(* IEC 61131-3 sources: POMIRTS_lab3/AS/Library_2/AsSafety, 3 files *)

(* ---- AsSafety.fun ---- *)
{REDUND_ERROR} FUNCTION_BLOCK safeRemoteControl (*Remote Control Function Block*)
	VAR_INPUT
		SafeLOGICID : UINT; (*SafeLOGIC ID*)
		Execute : BOOL; (*execution*)
		pCommandData : UDINT; (*pointer to command data*)
	END_VAR
	VAR_OUTPUT
		Done : BOOL; (*execution done*)
		Busy : BOOL; (*execution busy*)
		Error : BOOL; (*execution error*)
		StatusID : UINT; (*execution status: ERR_OK, ERR_FUB_BUSY, 0xXXXX = see help*)
		SafeLOGICStatus : RemoteControlStatusTypeV1; (*SafeLOGIC status*)
	END_VAR
	VAR
		i_state : UINT; (*internal variable*)
		i_result : UINT; (*internal variable*)
		i_tmp : UDINT; (*internal variable*)
		i_handle : UDINT; (*internal variable*)
	END_VAR
END_FUNCTION_BLOCK

{REDUND_ERROR} FUNCTION_BLOCK safeRemoteControl_V2 (*Remote Control Function Block*)
	VAR_INPUT
		SafeLOGICID : UINT; (*SafeLOGIC ID*)
		Execute : BOOL; (*execution*)
		pCommandData : UDINT; (*pointer to command data*)
	END_VAR
	VAR_OUTPUT
		Done : BOOL; (*execution done*)
		Busy : BOOL; (*execution busy*)
		Error : BOOL; (*execution error*)
		StatusID : UINT; (*execution status: ERR_OK, ERR_FUB_BUSY, 0xXXXX = see help*)
		SafeLOGICStatus : RemoteControlStatusTypeV2; (*SafeLOGIC status*)
	END_VAR
	VAR
		Internal : AsSafetyInternalType; (*internal variable*)
	END_VAR
END_FUNCTION_BLOCK

{REDUND_ERROR} FUNCTION_BLOCK safeDownloadApplication (*Download Application Function Block*)
	VAR_INPUT
		SafeLOGICID : UINT; (*SafeLOGIC ID*)
		Execute : BOOL; (*execution*)
		pCommandData : UDINT; (*pointer to command data*)
	END_VAR
	VAR_OUTPUT
		Done : BOOL; (*execution done*)
		Busy : BOOL; (*execution busy*)
		Error : BOOL; (*execution error*)
		StatusID : UINT; (*execution status: ERR_OK, ERR_FUB_BUSY, 0xXXXX = see help*)
		UnlockRequired : BOOL; (*unlock required*)
		ApplicationCRC : UDINT; (*application CRC*)
	END_VAR
	VAR
		i_state : UINT; (*internal variable*)
		i_result : UINT; (*internal variable*)
		i_tmp : UDINT; (*internal variable*)
		i_handle : UDINT; (*internal variable*)
	END_VAR
END_FUNCTION_BLOCK

{REDUND_ERROR} FUNCTION_BLOCK safeDownloadApplication_V2 (*Download Application Function Block*)
	VAR_INPUT
		SafeLOGICID : UINT; (*SafeLOGIC ID*)
		Execute : BOOL; (*execution*)
		pCommandData : UDINT; (*pointer to command data*)
	END_VAR
	VAR_OUTPUT
		Done : BOOL; (*execution done*)
		Busy : BOOL; (*execution busy*)
		Error : BOOL; (*execution error*)
		StatusID : UINT; (*execution status: ERR_OK, ERR_FUB_BUSY, 0xXXXX = see help*)
		UnlockRequired : BOOL; (*unlock required*)
		ApplicationCRC : UDINT; (*application CRC*)
	END_VAR
	VAR
		Internal : AsSafetyInternalType; (*internal variable*)
	END_VAR
END_FUNCTION_BLOCK

{REDUND_ERROR} FUNCTION_BLOCK safeDownloadData (*Download Data Function Block*)
	VAR_INPUT
		SafeLOGICID : UINT; (*SafeLOGIC ID*)
		Execute : BOOL; (*execution*)
		Type : UINT; (*type of data: safeDATA_TYPE_MAOP, safeDATA_TYPE_EXTMAOP,... *)
		pCommandData : UDINT; (*pointer to command data*)
	END_VAR
	VAR_OUTPUT
		Done : BOOL; (*execution done*)
		Busy : BOOL; (*execution busy*)
		Error : BOOL; (*execution error*)
		StatusID : UINT; (*execution status: ERR_OK, ERR_FUB_BUSY, 0xXXXX = see help*)
		UnlockRequired : BOOL; (*unlock required*)
		Timestamp : UDINT; (*timestamp from data*)
	END_VAR
	VAR
		i_state : UINT; (*internal variable*)
		i_result : UINT; (*internal variable*)
		i_tmp : UDINT; (*internal variable*)
		i_handle : UDINT; (*internal variable*)
	END_VAR
END_FUNCTION_BLOCK

{REDUND_ERROR} FUNCTION_BLOCK safeDownloadData_V2 (*Download Data Function Block*)
	VAR_INPUT
		SafeLOGICID : UINT; (*SafeLOGIC ID*)
		Execute : BOOL; (*execution*)
		Type : UINT; (*type of data: safeDATA_TYPE_MAOP, safeDATA_TYPE_EXTMAOP,... *)
		pCommandData : UDINT; (*pointer to command data*)
	END_VAR
	VAR_OUTPUT
		Done : BOOL; (*execution done*)
		Busy : BOOL; (*execution busy*)
		Error : BOOL; (*execution error*)
		StatusID : UINT; (*execution status: ERR_OK, ERR_FUB_BUSY, 0xXXXX = see help*)
		UnlockRequired : BOOL; (*unlock required*)
		Timestamp : UDINT; (*timestamp from data*)
	END_VAR
	VAR
		Internal : AsSafetyInternalType; (*internal variable*)
	END_VAR
END_FUNCTION_BLOCK

{REDUND_ERROR} FUNCTION_BLOCK safeConfigurationOnTarget (*Configuration On Target Function Block*)
	VAR_INPUT
		SafeLOGICID : UINT; (*SafeLOGIC ID*)
		Execute : BOOL; (*execution*)
		Type : UINT; (*type of data: safeDATA_TYPE_MAOP, safeDATA_TYPE_EXTMAOP,...*)
		pCommandData : UDINT; (*pointer to command data*)
	END_VAR
	VAR_OUTPUT
		Done : BOOL; (*execution done*)
		Busy : BOOL; (*execution busy*)
		Error : BOOL; (*execution error*)
		StatusID : UINT; (*execution status: ERR_OK, ERR_FUB_BUSY, 0xXXXX = see help*)
		Timestamp : UDINT; (*timestamp of data*)
	END_VAR
	VAR
		i_state : UINT; (*internal variable*)
		i_result : UINT; (*internal variable*)
		i_tmp : UDINT; (*internal variable*)
		i_handle : UDINT; (*internal variable*)
	END_VAR
END_FUNCTION_BLOCK

{REDUND_ERROR} FUNCTION_BLOCK safeConfigurationOnTarget_V2 (*Configuration On Target Function Block*)
	VAR_INPUT
		SafeLOGICID : UINT; (*SafeLOGIC ID*)
		Execute : BOOL; (*execution*)
		Type : UINT; (*type of data: safeDATA_TYPE_MAOP, safeDATA_TYPE_EXTMAOP,...*)
		pCommandData : UDINT; (*pointer to command data*)
	END_VAR
	VAR_OUTPUT
		Done : BOOL; (*execution done*)
		Busy : BOOL; (*execution busy*)
		Error : BOOL; (*execution error*)
		StatusID : UINT; (*execution status: ERR_OK, ERR_FUB_BUSY, 0xXXXX = see help*)
		Timestamp : UDINT; (*timestamp of data*)
	END_VAR
	VAR
		Internal : AsSafetyInternalType; (*internal variable*)
	END_VAR
END_FUNCTION_BLOCK

{REDUND_ERROR} FUNCTION safeLibraryVersion : UINT (*returns the actual library version*)
END_FUNCTION

{REDUND_ERROR} FUNCTION_BLOCK safeDownloadFile (*Download File Function Block*)
	VAR_INPUT
		SafeLOGICID : UINT; (*SafeLOGIC ID*)
		Execute : BOOL; (*execution*)
		pCommandData : UDINT; (*pointer to command data*)
	END_VAR
	VAR_OUTPUT
		Done : BOOL; (*execution done*)
		Busy : BOOL; (*execution busy*)
		Error : BOOL; (*execution error*)
		StatusID : UINT; (*execution status: ERR_OK, ERR_FUB_BUSY, 0xXXXX = see help*)
		UnlockRequired : BOOL; (*unlock required*)
		Timestamp : UDINT; (*timestamp from data*)
	END_VAR
	VAR
		Internal : AsSafetyInternalType; (*internal variable*)
	END_VAR
END_FUNCTION_BLOCK

{REDUND_ERROR} FUNCTION_BLOCK safeCheckTable (*Check Table Function Block*)
	VAR_INPUT
		Execute : BOOL; (*execution*)
		InstNr : USINT; (*instance number*)
		pUser : UDINT; (*user name*)
		Timestamp : UDINT; (*timestamp*)
		TableType : USINT; (*table type*)
		EntryCnt : UDINT; (*number of entries*)
		pTableHeader : UDINT; (*table header input*)
		pTableData : UDINT; (*table data input*)
		pTableHeaderOut : UDINT; (*table header output buffer*)
		pTableDataOut : UDINT; (*table data output buffer*)
		pFileDataOut : UDINT; (*file data output buffer*)
		AckData : USINT; (*1 .. acknowledge table data, 2 .. NOT acknowledge table data, abort FUB*)
	END_VAR
	VAR_OUTPUT
		Done : BOOL; (*execution done*)
		Busy : BOOL; (*execution busy*)
		Error : BOOL; (*execution error*)
		StatusID : UINT; (*execution status: ERR_OK, ERR_FUB_BUSY, 0xXXXX = see help*)
		CheckErrorCode : UDINT; (*table check error code*)
		CheckErrorLine : UDINT; (*table check error line*)
		CheckErrorColumn : UDINT; (*table check error column*)
		pCrcOut : UDINT; (*returns pointer to CRC data*)
		CrcCntOut : UDINT; (*returns number of CRCs*)
	END_VAR
	VAR
		i_step : UINT; (*internal*)
		i_tmp : UDINT; (*internal*)
		i_clean : BOOL; (*internal*)
	END_VAR
END_FUNCTION_BLOCK

{REDUND_ERROR} FUNCTION_BLOCK safeFileInfo (*File Info Function Block*)
	VAR_INPUT
		SafeLOGICID : UINT; (*SafeLOGIC ID*)
		Execute : BOOL; (*execution*)
		Type : UINT; (*type of data: safeDATA_TYPE_MAOP, safeDATA_TYPE_EXTMAOP,...*)
		pCommandData : UDINT; (*pointer to command data*)
	END_VAR
	VAR_OUTPUT
		Done : BOOL; (*execution done*)
		Busy : BOOL; (*execution busy*)
		Error : BOOL; (*execution error*)
		StatusID : UINT; (*execution status: ERR_OK, ERR_FUB_BUSY, 0xXXXX = see help*)
	END_VAR
	VAR
		Internal : AsSafetyInternalType; (*internal variable*)
	END_VAR
END_FUNCTION_BLOCK

{REDUND_ERROR} FUNCTION safeGetTableLength : UDINT (*Function returns size of table data*)
	VAR_INPUT
		TableType : USINT; (*table type*)
		EntryCnt : UDINT; (*number of entries*)
		pTableHeader : UDINT; (*pointer to table header*)
	END_VAR
END_FUNCTION

{REDUND_ERROR} FUNCTION_BLOCK safeGetDataLength (*Function Block returns size of download file*)
	VAR_INPUT
		Execute : BOOL; (*execution*)
		Type : UINT; (*type of data: safeDATA_TYPE_MAOP, safeDATA_TYPE_EXTMAOP,... *)
		pCommandData : UDINT; (*pointer to command data*)
	END_VAR
	VAR_OUTPUT
		Done : BOOL; (*execution done*)
		Busy : BOOL; (*execution busy*)
		Error : BOOL; (*execution error*)
		StatusID : UINT; (*execution status: ERR_OK, ERR_FUB_BUSY, 0xXXXX = see help*)
		Length : UDINT; (*calculated length of download file*)
	END_VAR
	VAR
		Internal : AsSafetyInternalType; (*internal variable*)
	END_VAR
END_FUNCTION_BLOCK

{REDUND_ERROR} FUNCTION_BLOCK safeCreateData (*Create Data Function Block*)
	VAR_INPUT
		SafeLOGICID : UINT; (*SafeLOGIC ID*)
		Execute : BOOL; (*execution*)
		Type : UINT; (*type of data: safeDATA_TYPE_MAOP, safeDATA_TYPE_EXTMAOP,... *)
		pCommandData : UDINT; (*pointer to command data*)
		FileDataOutLen : UDINT; (*size of buffer for file data*)
		pFileDataOut : UDINT; (*pointer to memory buffer for file data*)
	END_VAR
	VAR_OUTPUT
		Done : BOOL; (*execution done*)
		Busy : BOOL; (*execution busy*)
		Error : BOOL; (*execution error*)
		StatusID : UINT; (*execution status: ERR_OK, ERR_FUB_BUSY, 0xXXXX = see help*)
		UnlockRequired : BOOL; (*unlock required*)
		Timestamp : UDINT; (*timestamp from data*)
	END_VAR
	VAR
		Internal : AsSafetyInternalType; (*internal variable*)
	END_VAR
END_FUNCTION_BLOCK

{REDUND_ERROR} FUNCTION_BLOCK safeLogicInfo (*Remote Control Function Block*)
	VAR_INPUT
		SafeLOGICID : UINT; (*SafeLOGIC ID*)
		Execute : BOOL; (*execution*)
		Type : UINT; (*type of data: safeINFO_TYPE_PWD_INFO, safeINFO_TYPE_PWD_CHK, safeINFO_TYPE_UDID_INFO*)
		pCommandData : UDINT; (*pointer to command data*)
	END_VAR
	VAR_OUTPUT
		Done : BOOL; (*execution done*)
		Busy : BOOL; (*execution busy*)
		Error : BOOL; (*execution error*)
		StatusID : UINT; (*execution status: ERR_OK, ERR_FUB_BUSY, 0xXXXX = see help*)
	END_VAR
	VAR
		Internal : AsSafetyInternalType; (*internal variable*)
	END_VAR
END_FUNCTION_BLOCK

(* ---- AsSafety.typ ---- *)
TYPE
	FileReferenceType : 	STRUCT  (*file reference*)
		Device : STRING[80]; (*pointer to the device name*)
		File : STRING[80]; (*pointer to the file name*)
	END_STRUCT;
	AsSafetyInternalType : 	STRUCT  (*internal data type*)
		Clean : BOOL;
		State : UINT;
		Result : UINT;
		Tmp : UDINT;
		pThis : UDINT;
		pFcn : UDINT;
	END_STRUCT;
	SourceLocalDataTypeV1 : 	STRUCT  (*local data source type*)
		pFileData : UDINT; (*pointer to data buffer*)
		FileLength : UDINT; (*data length*)
	END_STRUCT;
	SourceLocalFileTypeV1 : 	STRUCT  (*local file source*)
		SourceFile : FileReferenceType; (*path to local file*)
	END_STRUCT;
	DataSourceTypeV1 : 	STRUCT  (*source data type*)
		Type : UINT; (*0 .. file upload from safeLOGIC, 1 .. local data buffer, 2 .. local file*)
		LocalData : SourceLocalDataTypeV1; (*arguments for local data*)
		LocalFile : SourceLocalFileTypeV1; (*arguments for local file*)
	END_STRUCT;
	InfoCmdPwdInfoTypeV1 : 	STRUCT  (*password info data from SafeLOGIC command structure*)
		Version : UINT; (*used version*)
		PasswordSet : BOOL; (*0 .. no password set, 1 .. password is set*)
	END_STRUCT;
	InfoCmdPwdChkTypeV1 : 	STRUCT  (*password check data from SafeLOGIC command structure*)
		Version : UINT; (*used version*)
		Password : STRING[16]; (*password for check*)
		PasswordEqual : BOOL; (*0 .. no password set, 1 .. password is set*)
	END_STRUCT;
	ConfigurationAddParaTypeV2 : 	STRUCT  (*additional parameter data from SafeLOGIC*)
		SADR : UINT; (*safety address*)
		ID : USINT; (*id*)
		pParaData : UDINT; (*pointer to additional parameter data*)
		Length : UDINT; (*size of parameter buffer*)
		LengthOut : UDINT; (*length of parameter*)
		CRC : UDINT; (*CRC*)
		Timestamp : UDINT; (*timestamp*)
	END_STRUCT;
	ConfigurationAddParaTypeV1 : 	STRUCT  (*additional parameter data from SafeLOGIC*)
		SADR : UINT; (*safety address*)
		ID : USINT; (*id*)
		pParaData : UDINT; (*pointer to additional parameter data*)
		Length : UDINT; (*size of parameter buffer*)
		CRC : UDINT; (*CRC*)
		Timestamp : UDINT; (*timestamp*)
	END_STRUCT;
	ConfigurationBitOptionsTypeV1 : 	STRUCT  (*bit machine options*)
		BitData : ARRAY[0..63]OF USINT; (*bit array*)
	END_STRUCT;
	ConfigurationCmdAddParaTypeV2 : 	STRUCT  (*additional parameter data from SafeLOGIC command structure*)
		Version : UINT; (*input data: used version*)
		Password : STRING[16]; (*input data: password*)
		pParaDataOutput : UDINT; (*input data: pointer to list of type ConfigurationAddParaTypeV2*)
		NumberParaSetsOutput : UINT; (*input data: number of available entries in pParaDataOutput*)
		NumberParaSetsOutputOut : UINT; (*return value: number of returned entries*)
		pBackupFile : UDINT; (*input data: 0 .. no backup, otherwise pointer to struct of type FileReferenceType *)
		pXmlOutputFile : UDINT; (*input data: 0 .. don't create XML output data, otherwise pointer to struct of type FileReferenceType*)
	END_STRUCT;
	ConfigurationCmdAddParaTypeV1 : 	STRUCT  (*additional parameter data from SafeLOGIC command structure*)
		Version : UINT; (*input data: used version*)
		Password : STRING[16]; (*input data: password*)
		pParaDataOutput : UDINT; (*return value: pointer to list of type ConfigurationAddParaTypeV1*)
		NumberParaSetsOutput : UINT; (*return value: number of returned entries*)
	END_STRUCT;
	ConfigurationCmdExtMaOpTypeV2 : 	STRUCT  (*extended machine options from SafeLOGIC command structure*)
		Version : UINT; (*input data: safeVERSION_R110*)
		Password : STRING[16]; (*input data: password*)
		pIntDataOutput : UDINT; (*input data: pointer to list of type ConfigurationIntOptionsTypeV1*)
		NumberIntOutput : UINT; (*input data: number of available entries in INT buffer*)
		NumberIntOutputOut : UINT; (*return value: number of returned INT data entries*)
		pUintDataOutput : UDINT; (*input data: pointer to list of type ConfigurationUintOptionsTypeV1*)
		NumberUintOutput : UINT; (*input data: number of available entries in UINT buffer*)
		NumberUintOutputOut : UINT; (*return value: number of returned UINT data entries*)
		pDintDataOutput : UDINT; (*input data: pointer to list of type ConfigurationDintOptionsTypeV1*)
		NumberDintOutput : UINT; (*input data: number of available DINT data entries*)
		NumberDintOutputOut : UINT; (*return value: number of returned DINT data entries*)
		pUdintDataOutput : UDINT; (*input data: pointer to list of type ConfigurationUdintOptionsTypeV1*)
		NumberUdintOutput : UINT; (*input data: number of available UDINT data entries*)
		NumberUdintOutputOut : UINT; (*return value: number of returned UDINT data entries*)
		pBackupFile : UDINT; (*input data: 0 .. no backup, otherwise pointer to struct of type FileReferenceType *)
		pXmlOutputFile : UDINT; (*input data: 0 .. don't create XML output data, otherwise pointer to struct of type FileReferenceType*)
	END_STRUCT;
	ConfigurationCmdExtMaOpTypeV1 : 	STRUCT  (*extended machine options from SafeLOGIC command structure*)
		Version : UINT; (*input data: safeVERSION_R107*)
		Password : STRING[16]; (*input data: password*)
		pIntDataOutput : UDINT; (*return value: pointer to list of type ConfigurationIntOptionsTypeV1*)
		NumberIntOutput : UINT; (*return value: number of returned INT data entries*)
		pUintDataOutput : UDINT; (*return value: pointer to list of type ConfigurationUintOptionsTypeV1*)
		NumberUintOutput : UINT; (*return value: number of returned UINT data entries*)
		pDintDataOutput : UDINT; (*return value: pointer to list of type ConfigurationDintOptionsTypeV1*)
		NumberDintOutput : UINT; (*return value: number of returned DINT data entries*)
		pUdintDataOutput : UDINT; (*return value: pointer to list of type ConfigurationUdintOptionsTypeV1*)
		NumberUdintOutput : UINT; (*return value: number of returned UDINT data entries*)
	END_STRUCT;
	ConfigurationCmdMaOpTypeV2 : 	STRUCT  (*machine options from SafeLOGIC command structure Version 2*)
		Version : UINT; (*input data: safeVERSION_R110*)
		Password : STRING[16]; (*input data: password*)
		pDeviceListOutput : UDINT; (*input data: pointer to device list buffer of type ConfigurationDeviceTypeV1*)
		NumberDevicesOutput : UINT; (*input data: number of available device entries in devices list buffer*)
		NumberDevicesOutputOut : UINT; (*return value: number of returned device entries*)
		pMachineOptionsOutput : UDINT; (*input data: pointer to bit machine options of type ConfigurationBitOptionsTypeV1*)
		pModuleFlagsOutput : UDINT; (*input data: pointer to module flags of type ConfigurationModuleFlagsTypeV1*)
		pBackupFile : UDINT; (*input data: 0 .. no backup, otherwise pointer to struct of type FileReferenceType *)
		pXmlOutputFile : UDINT; (*input data: 0 .. don't create XML output data, otherwise pointer to struct of type FileReferenceType*)
	END_STRUCT;
	ConfigurationCmdMaOpTypeV1 : 	STRUCT  (*machine options from SafeLOGIC command structure Version 1*)
		Version : UINT; (*input data: safeVERSION_R107*)
		Password : STRING[16]; (*input data: password*)
		pDeviceListOutput : UDINT; (*return value: pointer to device list of type ConfigurationDeviceTypeV1*)
		NumberDevicesOutput : UINT; (*return value: number of returned entries*)
		pMachineOptionsOutput : UDINT; (*return value: pointer to bit machine options of type ConfigurationBitOptionsTypeV1*)
		pModuleFlagsOutput : UDINT; (*return value: pointer to module flags of type ConfigurationModuleFlagsTypeV1*)
	END_STRUCT;
	ConfigurationCmdTableTypeV2 : 	STRUCT  (*table data from SafeLOGIC command structure*)
		Version : UINT; (*input data: safeVERSION_R110*)
		Password : STRING[16]; (*input data: password*)
		pTableDataOutput : UDINT; (*input data: pointer to list of type ConfigurationTableTypeV1*)
		NumberTablesOutput : UINT; (*input data: number of available entries in pTableDataOutput*)
		NumberTablesOutputOut : UINT; (*return value: number of returned table entries*)
		pBackupFile : UDINT; (*input data: 0 .. no backup, otherwise pointer to struct of type FileReferenceType *)
		pXmlOutputFile : UDINT; (*input data: 0 .. don't create XML output data, otherwise pointer to struct of type FileReferenceType*)
	END_STRUCT;
	ConfigurationCmdTableTypeV1 : 	STRUCT  (*table data from SafeLOGIC command structure*)
		Version : UINT; (*input data: safeVERSION_R107*)
		Password : STRING[16]; (*input data: password*)
		pTableDataOutput : UDINT; (*return value: pointer to list of type ConfigurationTableTypeV1*)
		NumberTablesOutput : UINT; (*return value: number of returned table entries*)
	END_STRUCT;
	FileInfoCmdTypeV1 : 	STRUCT  (*file info command structure*)
		Version : UINT; (*used version*)
		DataSource : DataSourceTypeV1; (*data source*)
		Timestamp : UDINT; (*timestamp*)
		pCrcs : UDINT; (*buffer for CRCs*)
		NumberOfCrcs : UINT; (*size of CRC buffer*)
		NumberOfCrcsOut : UINT; (*number of CRCs*)
	END_STRUCT;
	ConfigurationDeviceTypeV1 : 	STRUCT  (*safety device from SafeLOGIC*)
		SADR : UINT; (*safety address*)
		UDID : ARRAY[0..5]OF USINT; (*UDID*)
	END_STRUCT;
	ConfigurationDintOptionsTypeV1 : 	STRUCT  (*DINT machine options*)
		ID : UINT; (*id*)
		Value : DINT; (*value*)
	END_STRUCT;
	ConfigurationIntOptionsTypeV1 : 	STRUCT  (*INT machine options*)
		ID : UINT; (*id*)
		Value : INT; (*value*)
	END_STRUCT;
	ConfigurationModuleFlagsTypeV1 : 	STRUCT  (*module flags*)
		Optional : ARRAY[0..127]OF USINT; (*optional*)
		Startup : ARRAY[0..127]OF USINT; (*startup*)
		NotPresent : ARRAY[0..127]OF USINT; (*not present*)
	END_STRUCT;
	ConfigurationTableTypeV2 : 	STRUCT  (*table data for command struct V1*)
		ID : UINT; (*table id*)
		Type : USINT; (*table type*)
		NumberOfCRCs : UINT; (*input data: number of available entries in pCRCData*)
		NumberOfCRCsOut : UINT; (*return value: number of returned CRC entries*)
		pCRCData : UDINT; (*input data: pointer to table CRC buffer*)
	END_STRUCT;
	ConfigurationTableTypeV1 : 	STRUCT  (*table data for command struct V2*)
		ID : UINT; (*table id*)
		Type : USINT; (*table type*)
		NumberOfCRCs : UINT; (*return value: number of returned CRCs*)
		pCRCData : UDINT; (*return value: pointer to table CRC buffer*)
	END_STRUCT;
	ConfigurationUdintOptionsTypeV1 : 	STRUCT  (*UDINT machine options*)
		ID : UINT; (*id*)
		Value : UDINT; (*value*)
	END_STRUCT;
	ConfigurationUintOptionsTypeV1 : 	STRUCT  (*UINT machine options*)
		ID : UINT; (*id*)
		Value : UINT; (*value*)
	END_STRUCT;
	DownloadAcknExtMaOpTypeV1 : 	STRUCT  (*acknowledge extended machine options structure*)
		AcknIntOptions : ARRAY[0..63]OF BOOL; (*acknowledge INT*)
		AcknUintOptions : ARRAY[0..63]OF BOOL; (*acknowledge UINT*)
		AcknDintOptions : ARRAY[0..63]OF BOOL; (*acknowledge DINT*)
		AcknUdintOptions : ARRAY[0..63]OF BOOL; (*acknowledge UDINT*)
	END_STRUCT;
	DownloadAcknMaOpTypeV1 : 	STRUCT  (*acknowledge bit machine options structure*)
		AcknBitOptions : ARRAY[0..63]OF USINT; (*acknowledge bit*)
	END_STRUCT;
	DownloadAcknAddParaTypeV1 : 	STRUCT  (*acknowledge bit additional parameter*)
		AcknBitAddPara : ARRAY[0..63]OF USINT; (*acknowledge bit*)
	END_STRUCT;
	DownloadCmdAddParaTypeV2 : 	STRUCT  (*additional paramater command structure*)
		Version : UINT; (*input data: used version*)
		Password : STRING[16]; (*input data: password*)
		UDID_Low : UDINT; (*input data: UDID low*)
		UDID_High : UINT; (*input data: UDID high*)
		Unlock : USINT; (*input data: unlock data*)
		pParaListInput : UDINT; (*input data: pointer to additional parameter input data list of type DownloadAddParaTypeV1*)
		NumberParaSetsInput : UINT; (*input data: number of input parameter entries in pParaListInput*)
		pParaDataOutput : UDINT; (*input data: pointer to list of type ConfigurationAddParaTypeV2*)
		NumberParaSetsOutput : UINT; (*input data: number of available entries in pParaDataOutput*)
		NumberParaSetsOutputOut : UINT; (*return value: number of returned entries*)
		pBackupFile : UDINT; (*input data: 0 .. no backup, otherwise pointer to struct of type FileReferenceType *)
		pXmlOutputFile : UDINT; (*input data: 0 .. don't create XML output data, otherwise pointer to struct of type FileReferenceType*)
	END_STRUCT;
	DownloadCmdAddParaTypeV1 : 	STRUCT  (*additional paramater command structure*)
		Version : UINT; (*input data: used version*)
		Password : STRING[16]; (*input data: password*)
		UDID_Low : UDINT; (*input data: UDID low*)
		UDID_High : UINT; (*input data: UDID high*)
		Unlock : USINT; (*input data: unlock data*)
		pParaListInput : UDINT; (*input data: pointer to additional parameter input data list of type DownloadAddParaTypeV1*)
		NumberParaSetsInput : UINT; (*input data: number of input parameter entries in pParaListInput*)
		pParaDataOutput : UDINT; (*return value: pointer to list of type ConfigurationAddParaTypeV1*)
		NumberParaSetsOutput : UINT; (*return value: number of returned entries*)
	END_STRUCT;
	DownloadCmdApplicationTypeV1 : 	STRUCT  (*application command structure*)
		Version : UINT; (*used version*)
		Password : STRING[16]; (*password*)
		UDID_Low : UDINT; (*UDID low*)
		UDID_High : UINT; (*UDID high*)
		ApplicationID : UINT; (*application id*)
		Device : STRING[80]; (*device for file*)
		File : STRING[80]; (*file name*)
		Unlock : USINT; (*unlock application*)
	END_STRUCT;
	DownloadCmdExtMaOpTypeV2 : 	STRUCT  (*extended machine options command structure*)
		Version : UINT; (*input data: safeVERSION_R110*)
		Password : STRING[16]; (*input data: password*)
		UDID_Low : UDINT; (*input data: UDID low*)
		UDID_High : UINT; (*input data: UDID high*)
		Unlock : USINT; (*input data: unlock data*)
		pIntDataInput : UDINT; (*input data: pointer to INT input data list from type ConfigurationIntOptionsTypeV1*)
		NumberIntInput : UINT; (*input data: number of INT input entries in pIntDataInput*)
		pUintDataInput : UDINT; (*input data: pointer to UINT input data list from type ConfigurationUintOptionsTypeV1*)
		NumberUintInput : UINT; (*input data: number of UINT input entries in pUintDataInput*)
		pDintDataInput : UDINT; (*input data: pointer to DINT input data list from type ConfigurationDintOptionsTypeV1*)
		NumberDintInput : UINT; (*input data: number of DINT input entries in pDintDataInput*)
		pUdintDataInput : UDINT; (*input data: pointer to UDINT input data list from type ConfigurationUdintOptionsTypeV1*)
		NumberUdintInput : UINT; (*input data: number of UDINT input entries in pUdintDataInput*)
		pAcknMachineOptions : UDINT; (*input data: pointer to acknowledge information of type DownloadAcknMaOpTypeV1*)
		pIntDataOutput : UDINT; (*input data: pointer to list of type ConfigurationIntOptionsTypeV1*)
		NumberIntOutput : UINT; (*input data: number of available entries in INT buffer*)
		NumberIntOutputOut : UINT; (*return value: number of returned INT data entries*)
		pUintDataOutput : UDINT; (*input data: pointer to list of type ConfigurationUintOptionsTypeV1*)
		NumberUintOutput : UINT; (*input data: number of available entries in UINT buffer*)
		NumberUintOutputOut : UINT; (*return value: number of returned UINT data entries*)
		pDintDataOutput : UDINT; (*input data: pointer to list of type ConfigurationDintOptionsTypeV1*)
		NumberDintOutput : UINT; (*input data: number of available DINT data entries*)
		NumberDintOutputOut : UINT; (*return value: number of returned DINT data entries*)
		pUdintDataOutput : UDINT; (*input data: pointer to list of type ConfigurationUdintOptionsTypeV1*)
		NumberUdintOutput : UINT; (*input data: number of available UDINT data entries*)
		NumberUdintOutputOut : UINT; (*number of UDINT channels from SafeLOGIC*)
		pBackupFile : UDINT; (*input data: 0 .. no backup, otherwise pointer to struct of type FileReferenceType *)
		pXmlOutputFile : UDINT; (*input data: 0 .. don't create XML output data, otherwise pointer to struct of type FileReferenceType*)
	END_STRUCT;
	DownloadCmdExtMaOpTypeV1 : 	STRUCT  (*return value: number of returned UDINT data entries*)
		Version : UINT; (*input data: safeVERSION_R107*)
		Password : STRING[16]; (*input data: password*)
		UDID_Low : UDINT; (*input data: UDID low*)
		UDID_High : UINT; (*input data: UDID high*)
		Unlock : USINT; (*input data: unlock data*)
		pIntDataInput : UDINT; (*input data: pointer to INT input data list from type ConfigurationIntOptionsTypeV1*)
		NumberIntInput : UINT; (*input data: number of INT input entries in pIntDataInput*)
		pUintDataInput : UDINT; (*input data: pointer to UINT input data list from type ConfigurationUintOptionsTypeV1*)
		NumberUintInput : UINT; (*input data: number of UINT input entries in pUintDataInput*)
		pDintDataInput : UDINT; (*input data: pointer to DINT input data list from type ConfigurationDintOptionsTypeV1*)
		NumberDintInput : UINT; (*input data: number of DINT input entries in pDintDataInput*)
		pUdintDataInput : UDINT; (*input data: pointer to UDINT input data list from type ConfigurationUdintOptionsTypeV1*)
		NumberUdintInput : UINT; (*input data: number of UDINT input entries in pUdintDataInput*)
		pAcknMachineOptions : UDINT; (*input data: pointer to acknowledge information of type DownloadAcknMaOpTypeV1*)
		pIntDataOutput : UDINT; (*return value: pointer to list of type ConfigurationIntOptionsTypeV1*)
		NumberIntOutput : UINT; (*return value: number of returned INT data entries*)
		pUintDataOutput : UDINT; (*return value: pointer to list of type ConfigurationUintOptionsTypeV1*)
		NumberUintOutput : UINT; (*return value: number of returned UINT data entries*)
		pDintDataOutput : UDINT; (*return value: pointer to list of type ConfigurationDintOptionsTypeV1*)
		NumberDintOutput : UINT; (*return value: number of returned DINT data entries*)
		pUdintDataOutput : UDINT; (*return value: pointer to list of type ConfigurationUdintOptionsTypeV1*)
		NumberUdintOutput : UINT; (*return value: number of returned UDINT data entries*)
	END_STRUCT;
	DownloadCmdMaOpTypeV2 : 	STRUCT  (*machine options command structure*)
		Version : UINT; (*input data: safeVERSION_R110*)
		Password : STRING[16]; (*input data: password*)
		UDID_Low : UDINT; (*input data: UDID low from SafeLOGIC*)
		UDID_High : UINT; (*input data: UDID high from SafeLOGIC*)
		Unlock : USINT; (*input data: unlock data*)
		pDeviceListInput : UDINT; (*input data: pointer to input device list of type DownloadDeviceTypeV1*)
		NumberDevicesInput : UINT; (*input data: number of input devices*)
		pMachineOptionsInput : UDINT; (*input data: pointer to input bit machine options of type ConfigurationBitOptionsTypeV1*)
		pModuleFlagsInput : UDINT; (*input data: pointer to input module flags of type ConfigurationModuleFlagsTypeV1*)
		pAcknMachineOptions : UDINT; (*input data: pointer to acknowledge information of type DownloadAcknMaOpTypeV1*)
		pDeviceListOutput : UDINT; (*input data: pointer to device list buffer of type ConfigurationDeviceTypeV1*)
		NumberDevicesOutput : UINT; (*input data: number of available device entries in devices list buffer*)
		NumberDevicesOutputOut : UINT; (*return value: number of returned device entries*)
		pMachineOptionsOutput : UDINT; (*input data: pointer to bit machine options of type ConfigurationBitOptionsTypeV1*)
		pModuleFlagsOutput : UDINT; (*input data: pointer to module flags of type ConfigurationModuleFlagsTypeV1*)
		pBackupFile : UDINT; (*input data: 0 .. no backup, otherwise pointer to struct of type FileReferenceType *)
		pXmlOutputFile : UDINT; (*input data: 0 .. don't create XML output data, otherwise pointer to struct of type FileReferenceType*)
	END_STRUCT;
	DownloadCmdMaOpTypeV1 : 	STRUCT  (*machine options command structure*)
		Version : UINT; (*input data: safeVERSION_R107*)
		Password : STRING[16]; (*input data: password*)
		UDID_Low : UDINT; (*input data: UDID low from SafeLOGIC*)
		UDID_High : UINT; (*input data: UDID high from SafeLOGIC*)
		Unlock : USINT; (*input data: unlock data*)
		pDeviceListInput : UDINT; (*input data: pointer to input device list of type DownloadDeviceTypeV1*)
		NumberDevicesInput : UINT; (*input data: number of input devices*)
		pMachineOptionsInput : UDINT; (*input data: pointer to input bit machine options of type ConfigurationBitOptionsTypeV1*)
		pModuleFlagsInput : UDINT; (*input data: pointer to input module flags of type ConfigurationModuleFlagsTypeV1*)
		pAcknMachineOptions : UDINT; (*input data: pointer to acknowledge information of type DownloadAcknMaOpTypeV1*)
		pDeviceListOutput : UDINT; (*return value: pointer to device list of type ConfigurationDeviceTypeV1*)
		NumberDevicesOutput : UINT; (*return value: number of returned entries*)
		pMachineOptionsOutput : UDINT; (*return value: pointer to bit machine options of type ConfigurationBitOptionsTypeV1*)
		pModuleFlagsOutput : UDINT; (*return value: pointer to module flags of type ConfigurationModuleFlagsTypeV1*)
	END_STRUCT;
	DownloadCmdTableTypeV2 : 	STRUCT  (*table command structure*)
		Version : UINT; (*input data: safeVERSION_R110*)
		Password : STRING[16]; (*input data: password*)
		UDID_Low : UDINT; (*input data: UDID low*)
		UDID_High : UINT; (*input data: UDID high*)
		Unlock : USINT; (*input data: unlock data*)
		pTableDataInput : UDINT; (*input data: pointer to input table data list of type DownloadTableTypeV2*)
		NumberTablesInput : UINT; (*input data: number of input entries in pTableDataInput*)
		pTableDataOutput : UDINT; (*input data: pointer to list of type ConfigurationTableTypeV1*)
		NumberTablesOutput : UINT; (*input data: number of available entries in pTableDataOutput*)
		NumberTablesOutputOut : UINT; (*return value: number of returned table entries*)
		pBackupFile : UDINT; (*input data: 0 .. no backup, otherwise pointer to struct of type FileReferenceType *)
		pXmlOutputFile : UDINT; (*input data: 0 .. don't create XML output data, otherwise pointer to struct of type FileReferenceType*)
	END_STRUCT;
	DownloadCmdTableTypeV1 : 	STRUCT  (*table command structure*)
		Version : UINT; (*input data: safeVERSION_R107*)
		Password : STRING[16]; (*input data: password*)
		UDID_Low : UDINT; (*input data: UDID low*)
		UDID_High : UINT; (*input data: UDID high*)
		Unlock : USINT; (*input data: unlock data*)
		pTableDataInput : UDINT; (*input data: pointer to input table data list of type DownloadTableTypeV1*)
		NumberTablesInput : UINT; (*input data: number of input entries in pTableDataInput*)
		pTableDataOutput : UDINT; (*return value: pointer to list of type ConfigurationTableTypeV1*)
		NumberTablesOutput : UINT; (*return value: number of returned table entries*)
	END_STRUCT;
	DownloadCmdFileTypeV1 : 	STRUCT  (*file command structure*)
		Version : UINT; (*used version*)
		Password : STRING[16]; (*password*)
		UDID_Low : UDINT; (*UDID low*)
		UDID_High : UINT; (*UDID high*)
		Unlock : USINT; (*unlock data*)
		DataSource : DataSourceTypeV1; (*local data or local file available, file upload from safeLOGIC not available*)
		pCrcs : UDINT; (*pointer to CRC data buffer*)
		NumberOfCrcs : UINT; (*size of CRC data Buffer*)
		NumberOfCrcsOut : UINT; (*number of CRCs*)
	END_STRUCT;
	DownloadAddParaTypeV1 : 	STRUCT  (*additional parameter data*)
		SADR : UINT; (*safety address*)
		ID : USINT; (*id*)
		pParaData : UDINT; (*pointer to additional parameter data*)
		Length : UDINT; (*length*)
		pAcknAddPara : UDINT; (*pointer to acknowledge information*)
	END_STRUCT;
	DownloadDeviceTypeV1 : 	STRUCT  (*safety device*)
		SADR : UINT; (*safety address*)
		UDID_Low : UDINT; (*UDID low*)
		UDID_High : UINT; (*UDID high*)
	END_STRUCT;
	DownloadTableTypeV1 : 	STRUCT  (*table data*)
		Device : STRING[80]; (*device for file*)
		File : STRING[80]; (*file name*)
	END_STRUCT;
	DownloadTableTypeV2 : 	STRUCT  (*table data*)
		Type : UINT; (*safeTABLE_FILE_TYPE .. use Device / File, safeTABLE_DATA_TYPE .. use pData / DataLen*)
		Device : STRING[80]; (*device for file*)
		File : STRING[80]; (*file name*)
		pData : UDINT; (*pointer to table data *)
		DataLen : UDINT; (*length of table data*)
	END_STRUCT;
	RemoteControlCmdTypeV1 : 	STRUCT  (*remote control command structure*)
		Version : UINT; (*used version*)
		Command : UINT; (*command*)
		Number : UINT; (*actual number*)
		Data : UINT; (*data*)
		Password : STRING[16]; (*password*)
		NewPassword : STRING[16]; (*new password*)
	END_STRUCT;
	RemoteControlStatusTypeV1 : 	STRUCT  (*remote control status from SafeLOGIC*)
		Command : UINT; (*last received command*)
		Number : UINT; (*running number of last received command*)
		Status : UINT; (*status of command*)
		State : UINT; (*state of the last ENTER command*)
		EnterData : UINT; (*last received ENTER command that was correct executed*)
		EnterNumber : UINT; (*running number of the last received ENTER command*)
		EnterExecuteStatus : UINT; (*state of the last received ENTER command*)
		SafeOSState : USINT; (*status of the safety application*)
		SafeKEYChanged : USINT; (*SafeKEY has been exchanged*)
		LedTestActive : USINT; (*LED test active*)
		Scanning : USINT; (*module scan active*)
		openSAFETYstate : USINT; (*status of openSAFETY stack*)
		FailSafe : USINT; (*Fail-Safe status*)
		NumberOfMissingModules : UINT; (*number of missing modules*)
		NumberOfUDIDMismatches : UINT; (*number of mismatched modules*)
		NumberOfDifferentFirmware : UINT; (*number of modules with different firmware*)
		SADR : ARRAY[0..100]OF UINT; (*safety address array*)
		MissingModules : ARRAY[0..15]OF USINT; (*missing modules array*)
		UDIDMismatches : ARRAY[0..15]OF USINT; (*udid mismatch array*)
		DifferentFirmware : ARRAY[0..15]OF USINT; (*different firmware array*)
	END_STRUCT;
	RemoteControlStatusTypeV2 : 	STRUCT  (*remote control status from SafeLOGIC*)
		Command : UINT; (*last received command*)
		Number : UINT; (*running number of last received command*)
		Status : UINT; (*status of command*)
		State : UINT; (*state of the last ENTER command*)
		EnterData : UINT; (*last received ENTER command that was correct executed*)
		EnterNumber : UINT; (*running number of the last received ENTER command*)
		EnterExecuteStatus : UINT; (*state of the last received ENTER command*)
		SafeOSState : USINT; (*status of the safety application*)
		SafeKEYChanged : USINT; (*SafeKEY has been exchanged*)
		LedTestActive : USINT; (*LED test active*)
		Scanning : USINT; (*module scan active*)
		openSAFETYstate : USINT; (*status of openSAFETY stack*)
		FailSafe : USINT; (*Fail-Safe status*)
		NumberOfMissingModules : UINT; (*number of missing modules*)
		NumberOfUDIDMismatches : UINT; (*number of mismatched modules*)
		NumberOfDifferentFirmware : UINT; (*number of modules with different firmware*)
		SADR : ARRAY[0..299]OF UINT; (*safety address array*)
		MissingModules : ARRAY[0..39]OF USINT; (*missing modules array*)
		UDIDMismatches : ARRAY[0..39]OF USINT; (*udid mismatch array*)
		DifferentFirmware : ARRAY[0..39]OF USINT; (*different firmware array*)
		NumberOfConfiguredModules : UINT; (*number of configured modules*)
		SetupModeActive : USINT; (*setup mode active*)
		ProjectPresent : USINT;	(*project present*)
		PasswordSet : USINT; (*password set*)
		IsSL81xx : USINT; (*SCM is part of SL81xx*)
		IsSCMar : USINT; (*SCM is part of SCMar*)
		SetupModeSupported : USINT; (*setup mode is supported*)
	END_STRUCT;
	TableHeaderATypeV1 : 	STRUCT  (*header struct for table type A version 1*)
		xTol : DINT;
		yTol : DINT;
	END_STRUCT;
	TableEntryATypeV1 : 	STRUCT  (*entry struct for table type A version 1*)
		xVal : DINT;
		yVal : DINT;
		resVal : USINT;
	END_STRUCT;
	TableEntryBTypeV1 : 	STRUCT  (*entry struct for table type B version 1*)
		xVal : DINT;
		yVal : DINT;
		zVal : DINT;
		resVal : DINT;
	END_STRUCT;
	TableEntryCTypeV1 : 	STRUCT  (*entry struct for table type C version 1*)
		Zone : UINT;
		Position : UINT;
		Dimension : UINT;
	END_STRUCT;
	TableHeaderDTypeV1 : 	STRUCT  (*header struct for table type A version 1*)
		Surveillance : BYTE;
	END_STRUCT;
	TableEntryDTypeV1 : 	STRUCT  (*entry struct for table type D version 1*)
		Object : UINT;
		Type : UINT;
		MinimumBeam : UINT;
		MaximumBeam : UINT;
		Dimension : UINT;
		DimensionTolerance : UINT;
	END_STRUCT;
	TableHeaderETypeV1 : 	STRUCT  (*header struct for table type E version 1*)
		xDim : INT;
		yDim : INT;
	END_STRUCT;
	TableEntryETypeV1 : 	STRUCT  (*entry struct for table type D version 1*)
		Entry : DINT;
	END_STRUCT;
	TableEntrySTypeV1 : 	STRUCT  (*entry struct for table type S version 1*)
		LinkTargetObjectID : DINT;
		LinkTargetAxisType : DINT;
		LinkSourceObjectID : DINT;
		LinkSourceAxisType : DINT;
		LinkFactorNum : DINT;
		LinkFactorDenom : DINT;
	END_STRUCT;
	TableHeaderTTypeV1 : 	STRUCT  (*header struct for table type T version 1*)
		NumberOfActiveAxes : DINT; (*number of active axes*)
	END_STRUCT;
	TableEntryTTypeV1 : 	STRUCT  (*entry struct for table type T version 1*)
		KinObjID : DINT;
		KinObjType : DINT;
		KinObjTransX : DINT;
		KinObjTransY : DINT;
		KinObjTransZ : DINT;
		KinObjRotAngle1 : DINT;
		KinObjRotAngle2 : DINT;
		KinObjRotAngle3 : DINT;
		KinObjRotaryAxisDecRamp : DINT;
		KinObjRotaryAxisMaxAcc : DINT;
		KinObjLinearAxisDecRamp : DINT;
		KinObjLinearAxisMaxAcc : DINT;
	END_STRUCT;
	TableHeaderTTypeV2 : 	STRUCT  (*header struct for table type T version 2*)
		NumberOfTableObjects : UINT;
		VersionNumber : UINT;
		NumberOfActiveAxes : DINT;
	END_STRUCT;
	TableEntryTTypeV2 : 	STRUCT  (*entry struct for table type T version 2*)
		KinObjID : DINT;
		KinObjType : DINT;
		KinObjTransX : DINT;
		KinObjTransY : DINT;
		KinObjTransZ : DINT;
		KinObjRotAngle1 : DINT;
		KinObjRotAngle2 : DINT;
		KinObjRotAngle3 : DINT;
		KinObjRotaryAxisDecRamp : DINT;
		KinObjRotaryAxisMaxAcc : DINT;
		KinObjLinearAxisDecRamp : DINT;
		KinObjLinearAxisMaxAcc : DINT;
		KinObjActivateWireFrameModel : DINT;
		KinObjDistanceToBndElements : DINT;
	END_STRUCT;
	TableHeaderTTypeV3 : 	STRUCT  (*header struct for table type T version 3*)
		NumberOfTableObjects : UINT;
		VersionNumber : UINT;
		NumberOfActiveAxes : DINT;
	END_STRUCT;
	TableEntryTTypeV3 : 	STRUCT  (*entry struct for table type T version 3*)
		KinObjID : DINT;
		KinObjType : DINT;
		KinObjTransX : DINT;
		KinObjTransY : DINT;
		KinObjTransZ : DINT;
		KinObjRotAngle1 : DINT;
		KinObjRotAngle2 : DINT;
		KinObjRotAngle3 : DINT;
		KinObjRotaryAxisDecRamp : DINT;
		KinObjRotaryAxisMaxAcc : DINT;
		KinObjLinearAxisDecRamp : DINT;
		KinObjLinearAxisMaxAcc : DINT;
		KinObjActivateWireFrameModel : DINT;
		KinObjDistanceToBndElements : DINT;
	END_STRUCT;
	TableEntryUTypeV1 : 	STRUCT  (*entry struct for table type U version 1*)
		SpaceID : DINT;
		SpaceType : DINT;
		SpaceTransX : DINT;
		SpaceTransY : DINT;
		SpaceTransZ : DINT;
		SpaceRotAngle1 : DINT;
		SpaceRotAngle2 : DINT;
		SpaceRotAngle3 : DINT;
		SpaceDimensionX : DINT;
		SpaceDimensionY : DINT;
		SpaceDimensionZ : DINT;
	END_STRUCT;
	TableEntryVTypeV1 : 	STRUCT  (*entry struct for table type V version 1*)
		SpaceID : DINT;
		SpaceType : DINT;
		KinObjID : DINT;
		KinObjJointAxisType : DINT;
		SpaceMaxLimit : DINT;
		SpaceMinLimit : DINT;
	END_STRUCT;
	TableEntryWTypeV1 : 	STRUCT  (* entry struct for table type W version 1*)
		OrientID : DINT;
		OrientType : DINT;
		OrientTransX_RotAngle1 : DINT;
		OrientTransY_RotAngle2 : DINT;
		OrientTransZ_RotAngle3 : DINT;
	END_STRUCT;
END_TYPE

(* ---- AsSafety.var ---- *)
VAR CONSTANT
	safeVERSION_R107 : UINT := 16#107; (*safety release version - 1.7*)
	safeVERSION_R110 : UINT := 16#110; (*safety release version - 1.10*)
	safeDATA_TYPE_MAOP : UINT := 16#100; (*download type for machine options *)
	safeDATA_TYPE_EXTMAOP : UINT := 16#200; (*download type for extended machine options *)
	safeDATA_TYPE_TABLE : UINT := 16#300; (*download type for table objects *)
	safeDATA_TYPE_ADDPARA : UINT := 16#400; (*download type for additional parameter*)
	safeDATA_TYPE_APPLICATION : UINT := 16#1200; (*type for restore*)
	safeINFO_TYPE_PWD_INFO : UINT := 1; (*SL info type for password info*)
	safeINFO_TYPE_PWD_CHK : UINT := 2; (*SL info type for password check*)
	safeTABLE_FILE_TYPE : UINT := 16#0000; (*reference to table file*)
	safeTABLE_DATA_TYPE : UINT := 16#0001; (*pointer to table data*)
	safeSRC_TYPE_UPLOAD_FILE : UINT := 0; (*file upload from SafeLOGIC*)
	safeSRC_TYPE_LOCAL_DATA : UINT := 1; (*local data from memory buffer*)
	safeSRC_TYPE_LOCAL_FILE : UINT := 2; (*local data from file*)
	safeCMD_ENTER : UINT := 16#100; (*enter command*)
	safeCMD_STATUS : UINT := 16#200; (*status command*)
	safeCMD_STATUS_SL : UINT := 16#0000; (*read back status*)
	safeCMD_N_UDID_ACKN : UINT := 16#20; (*acknowledge N modules*)
	safeCMD_4_UDID_ACKN : UINT := 16#30; (*acknowledge 4 modules*)
	safeCMD_3_UDID_ACKN : UINT := 16#40; (*acknowledge 3 modules*)
	safeCMD_2_UDID_ACKN : UINT := 16#50; (*acknowledge 2 modules*)
	safeCMD_1_UDID_ACKN : UINT := 16#60; (*acknowledge 1 module*)
	safeCMD_FW_ACKN : UINT := 16#100; (*acknowledge firmware*)
	safeCMD_SK_XCHG : UINT := 16#200; (*acknowledge SafeKEY*)
	safeCMD_TEST : UINT := 16#1000; (*LED test*)
	safeCMD_SCAN : UINT := 16#2000; (*scan*)
	safeCMD_SK_PW : UINT := 16#5000; (*change password*)
	safeCMD_SK_FORMAT : UINT := 16#6000; (*format SafeKEY*)
	safeCMD_RESET : UINT := 16#7000; (*reset SafeLOGIC*)
	safeCMD_CLEAR_DATA : UINT := 16#8000; (*clear additonal downloaded data*)
	safeCMD_SETUP_MODE_ACT : UINT := 16#9000; (*activate setup mode*)
	safeCMD_SETUP_MODE_DEACT : UINT := 16#9100; (*deactivate setup mode*)
	safeCMD_VERSION_INFO : UINT := 16#F000; (*remote version info*)
	safeRET_NO_TIMESTAMP : UDINT := 16#FFFFFFFF; (*no timestamp available*)
	safeERR_VERSION : UINT := 36100; (*error wrong version for command structure*)
	safeERR_PW_LENGTH : UINT := 36101; (*error wrong password length*)
	safeERR_UDID : UINT := 36102; (*error no UDID*)
	safeERR_ALLOC_MEM : UINT := 36103; (*error allocating memory*)
	safeERR_INTERNAL_ERROR : UINT := 36104; (*internal error*)
	safeERR_TIMEOUT : UINT := 36105; (*error connection timeout*)
	safeERR_RC_CMD : UINT := 36106; (*error wrong command*)
	safeERR_RC_ENTER_DATA : UINT := 36107; (*error wrong data for ENTER command*)
	safeERR_RC_ENTER_PW : UINT := 36108; (*error no password for command*)
	safeERR_RC_ENTER_SK_PW : UINT := 36109; (*error no new password for command*)
	safeERR_RC_STATUS_DATA : UINT := 36110; (*error wrong data for STATUS command*)
	safeERR_RC_DATA_LENGTH : UINT := 36111; (*error worng length for status data*)
	safeERR_DL_NO_PASSWORD : UINT := 36112; (*error no password for download*)
	safeERR_DL_PROTOCOL : UINT := 36113; (*error protocol version for download*)
	safeERR_DL_FILE_OPEN : UINT := 36114; (*error file open*)
	safeERR_DL_FILE_INVALID : UINT := 36115; (*error file invalid*)
	safeERR_DL_FILE_TOO_BIG : UINT := 36116; (*error file too big*)
	safeERR_DL_WRITE : UINT := 36117; (*error write*)
	safeERR_DL_STREAM : UINT := 36118; (*error stream*)
	safeERR_DL_CHECKSUM : UINT := 36119; (*error checksum*)
	safeERR_DL_UDID : UINT := 36120; (*error UDID doesn't match*)
	safeERR_DL_WRONG_FILE_SIZE : UINT := 36121; (*error wrong file size*)
	safeERR_DL_NO_RIGHTS_TO_WRITE : UINT := 36122; (*error wrong password*)
	safeERR_DL_UNLOCK_FILE_INFO : UINT := 36123; (*error file info*)
	safeERR_DL_UNLOCK_READ : UINT := 36124; (*error unlock read*)
	safeERR_DL_UNLOCK_WRITE : UINT := 36125; (*error unlock write*)
	safeERR_DL_STATIC_UNLOCK : UINT := 36126; (*error static unlock*)
	safeERR_DL_COMPARE_FAILED : UINT := 36127; (*error data compare failed*)
	safeERR_DLDATA_TYPE_ERR : UINT := 36128; (*error data type for download*)
	safeERR_DLDATA_ERR_DATA : UINT := 36129; (*error data for download*)
	safeERR_COT_TYPE_ERR : UINT := 36130; (*error data type for upload*)
	safeERR_COT_READING_FILE : UINT := 36131; (*error reading file*)
	safeERR_BUFFER_NULL : UINT := 36132; (*required input buffer is NULL*)
	safeERR_BUFFER_TOO_SMALL : UINT := 36133; (*required input buffer is too small*)
	safeERR_FILE_EMPTY : UINT := 36134; (*file is empty or does not exist on SL/SLX*)
	safeERR_FI_TYPE_ERR : UINT := 36135; (*error data type for getting file info*)
	safeERR_SLINFO_TYPE_ERR : UINT := 36136; (*error data type for SL info*)
	safeERR_SLINFO_RET_ERR : UINT := 36137; (*remote command returns error*)
	safeERR_COT_PWD_ERR : UINT := 36138; (*wrong password for configuration on target command*)
	safeERR_TC_INV_TABTYPE : UINT := 36180; (*invalid table type*)
	safeERR_TC_INV_INST : UINT := 36181; (*invalid table instance*)
	safeERR_TC_INV_INPUT_PTR : UINT := 36182; (*invalid input pointer*)
	safeERR_TC_INV_TAB_LEN : UINT := 36183; (*invalid table length*)
	safeERR_TC_INV_USER : UINT := 36184; (*invalid user name*)
	safeERR_TC_TYPE_CPY_FCT : UINT := 36185; (*no copy function for table type*)
	safeWRN_TC_WAIT_FOR_ACK : UINT := 36191; (*wait for acknowledge of tables*)
	safeERR_TC_CHECK_FAILED : UINT := 36186; (*table check failed*)
	safeERR_TC_EXTRACT_FAILED : UINT := 36187; (*extraction of output table data failed*)
	safeERR_TC_LOCK_FAILED : UINT := 36188; (*table lock failed*)
	safeERR_TC_ACK_SET : UINT := 36189; (*AckData is already set*)
	safeERR_TC_INVALID_STEP : UINT := 36190; (*invalid step in table check*)
END_VAR
